Fanuc KAREL source: kt00741.KL

PROGRAM KT00741
%STACKSIZE=65535
%PRIORITY=65535
%NOLOCKGROUP
VAR
ARG : ARRAY[4] OF SHORT
OUT : INTEGER
BEGIN
-- UNSAFE_SOURCE_IR line 7: OUT = native_s16_value(ARG)
END KT00741
